(* IEC 61131-3 sources: Test-Git_ESME26/TestProgettoESME_26.fbsproj/PacDriveLib Migration/Motion/Control/Brake, 3 files *)

(* ---- FB_BrakeCouplingTime.fb.st ---- *)
FUNCTION_BLOCK FB_BrakeCouplingTime IMPLEMENTS SE_Async.IF_Async
VAR
	xDone_loc          : BOOL;
	ifBrake_loc        : DDI.IF_Brake;
	tBrakeCouplingTemp : TIME := T#500MS;
END_VAR

(* ---- FB_BrakeDisconnectionTime.fb.st ---- *)
FUNCTION_BLOCK FB_BrakeDisconnectionTime IMPLEMENTS SE_Async.IF_Async
VAR
	xDone_loc            : BOOL;
	ifBrake_loc          : DDI.IF_Brake;
	tBrakeDisconnectTemp : TIME := T#500MS;
END_VAR

(* ---- FB_BrakeReleaseSet.fb.st ---- *)
FUNCTION_BLOCK INTERNAL FB_BrakeReleaseSet IMPLEMENTS SE_Async.IF_Async
VAR
	ifBrake_loc           : DDI.IF_Brake;
	xDone_loc             : BOOL;
	xRelease_loc          : BOOL;
END_VAR
